(* IEC 61131-3 sources: plc-st-coding-agent/progress/evidence/f14_v14_remaining_20261113/jobs/codex_minimax-m27 (part 2) *)

(* ---- public-hard-01.raw_candidate_02.st ---- *)
FUNCTION_BLOCK MaterialProportioning
VAR_INPUT
    estop           : BOOL;          // Emergency stop signal (FALSE = stopped)
    opeMode         : BOOL;          // Operation mode (FALSE = manual, TRUE = automatic)
    valveAStart     : BOOL;          // Valve A start button
    valveBStart     : BOOL;          // Valve B start button
    valveCStart     : BOOL;          // Valve C start button
    valveDStart     : BOOL;          // Valve D start button
    mixMotorStart   : BOOL;          // Mixing motor start button
    autoStart       : BOOL;          // Automatic start button
    processMode     : BOOL;          // Process mode (FALSE = simple, TRUE = with C)
    levelSensor     : INT;           // Liquid level sensor (cm)
    mixMotorComplete: BOOL;          // Mixing complete signal
END_VAR
VAR_OUTPUT
    valveARun       : BOOL;          // Valve A run command
    valveBRun       : BOOL;          // Valve B run command
    valveCRun       : BOOL;          // Valve C run command
    valveDRun       : BOOL;          // Valve D run command
    mixMotorRun     : BOOL;          // Mixing motor run command
END_VAR
VAR
    // Rising edge detection for manual toggle buttons
    tmp_autoStart        : R_TRIG;
    tmp_valveAStart      : R_TRIG;
    tmp_valveBStart      : R_TRIG;
    tmp_valveCStart      : R_TRIG;
    tmp_valveDStart      : R_TRIG;
    tmp_mixMotorStart    : R_TRIG;

    // Automatic mode state machine
    tmp_autoState   : INT;           // 0=idle, 1=fillA, 2=fillB, 3=fillC, 4=mix, 5=drain, 6=done

    // Manual mode toggle states
    tmp_manualValveA    : BOOL;
    tmp_manualValveB    : BOOL;
    tmp_manualValveC    : BOOL;
    tmp_manualValveD    : BOOL;
    tmp_manualMixMotor  : BOOL;

    // Process complete flag for automatic mode
    tmp_autoComplete    : BOOL;
END_VAR

(* ENGINEERING_CONTRACT
================================================================================
Output          | Activation                  | Retention      | Reset
----------------|------------------------------|----------------|-------------------------
valveARun       | Manual: rising valveAStart   | Hold toggle    | estop, opeMode, auto step
                | Auto: state=1, level<50      |                |
PUB001, PUB002, PUB003, PUB004, PUB005, PUB006, PUB007, PUB008
----------------|------------------------------|----------------|-------------------------
valveBRun       | Auto: state=2, level<80      | Hold until 80cm| estop, opeMode, auto step
                |                              |                |
PUB003, PUB004, PUB006, PUB007, PUB008
----------------|------------------------------|----------------|-------------------------
valveCRun       | Auto: state=3, level<100     | Hold until 100cm| estop, opeMode, auto step
                | (processMode=true only)      |                |
PUB003, PUB004, PUB006, PUB007, PUB008
----------------|------------------------------|----------------|-------------------------
valveDRun       | Auto: mixMotorComplete       | Hold until reset| estop, opeMode, autoStart
                |                              |                |
PUB007, PUB008, PUB011, PUB012, PUB013, PUB014, PUB015
----------------|------------------------------|----------------|-------------------------
mixMotorRun     | Auto: state=4                | Hold until complete| estop, opeMode, autoStart
                | Manual: rising mixMotorStart |                |
PUB007, PUB008, PUB011, PUB012, PUB013, PUB014, PUB015
================================================================================
Priority: estop > manual/automatic mode switch > same-scan state updates
Boundary: levelSensor thresholds at 50cm, 80cm, 100cm (>= comparisons)
================================================================================
*)

(* CONTRACT_RULES [] *)

// Detect rising edges for toggle buttons
tmp_autoStart(CLK := autoStart);
tmp_valveAStart(CLK := valveAStart);
tmp_valveBStart(CLK := valveBStart);
tmp_valveCStart(CLK := valveCStart);
tmp_valveDStart(CLK := valveDStart);
tmp_mixMotorStart(CLK := mixMotorStart);

// Emergency stop: all equipment OFF immediately
IF NOT estop THEN
    valveARun := FALSE;
    valveBRun := FALSE;
    valveCRun := FALSE;
    valveDRun := FALSE;
    mixMotorRun := FALSE;
    tmp_autoState := 0;
    tmp_autoComplete := FALSE;
    tmp_manualValveA := FALSE;
    tmp_manualValveB := FALSE;
    tmp_manualValveC := FALSE;
    tmp_manualValveD := FALSE;
    tmp_manualMixMotor := FALSE;
    RETURN;
END_IF;

// Mode selection
IF opeMode THEN
    // AUTOMATIC MODE
    // Rising edge of autoStart initiates process
    IF tmp_autoStart.Q AND tmp_autoState = 0 THEN
        tmp_autoState := 1;
        tmp_autoComplete := FALSE;
    END_IF;

    // State machine execution
    CASE tmp_autoState OF
        0:  // Idle - all off
            valveARun := FALSE;
            valveBRun := FALSE;
            valveCRun := FALSE;
            valveDRun := FALSE;
            mixMotorRun := FALSE;

        1:  // Fill with valve A until level >= 50cm
            valveARun := TRUE;
            valveBRun := FALSE;
            valveCRun := FALSE;
            valveDRun := FALSE;
            mixMotorRun := FALSE;
            IF levelSensor >= 50 THEN
                valveARun := FALSE;
                tmp_autoState := 2;
            END_IF;

        2:  // Fill with valve B until level >= 80cm
            valveARun := FALSE;
            valveBRun := TRUE;
            valveCRun := FALSE;
            valveDRun := FALSE;
            mixMotorRun := FALSE;
            IF levelSensor >= 80 THEN
                valveBRun := FALSE;
                // Check processMode to determine next state
                IF processMode THEN
                    tmp_autoState := 3;  // Go to valve C
                ELSE
                    tmp_autoState := 4;  // Go directly to mixing
                END_IF;
            END_IF;

        3:  // Fill with valve C (processMode=true) until level >= 100cm
            valveARun := FALSE;
            valveBRun := FALSE;
            valveCRun := TRUE;
            valveDRun := FALSE;
            mixMotorRun := FALSE;
            IF levelSensor >= 100 THEN
                valveCRun := FALSE;
                tmp_autoState := 4;
            END_IF;

        4:  // Mixing until mixMotorComplete signal
            valveARun := FALSE;
            valveBRun := FALSE;
            valveCRun := FALSE;
            valveDRun := FALSE;
            mixMotorRun := TRUE;
            IF mixMotorComplete THEN
                mixMotorRun := FALSE;
                tmp_autoState := 5;
            END_IF;

        5:  // Open valve D to drain
            valveARun := FALSE;
            valveBRun := FALSE;
            valveCRun := FALSE;
            valveDRun := TRUE;
            mixMotorRun := FALSE;
            tmp_autoComplete := TRUE;
            tmp_autoState := 6;

        6:  // Process complete - valve D remains open until reset
            valveARun := FALSE;
            valveBRun := FALSE;
            valveCRun := FALSE;
            valveDRun := TRUE;
            mixMotorRun := FALSE;
            // Wait for autoStart to reset
            IF tmp_autoStart.Q THEN
                tmp_autoState := 0;
                tmp_autoComplete := FALSE;
            END_IF;
    END_CASE;

ELSE
    // MANUAL MODE
    // Reset automatic state when switching to manual
    tmp_autoState := 0;
    tmp_autoComplete := FALSE;

    // Toggle valve A
    IF tmp_valveAStart.Q THEN
        tmp_manualValveA := NOT tmp_manualValveA;
    END_IF;

    // Toggle valve B
    IF tmp_valveBStart.Q THEN
        tmp_manualValveB := NOT tmp_manualValveB;
    END_IF;

    // Toggle valve C
    IF tmp_valveCStart.Q THEN
        tmp_manualValveC := NOT tmp_manualValveC;
    END_IF;

    // Toggle valve D
    IF tmp_valveDStart.Q THEN
        tmp_manualValveD := NOT tmp_manualValveD;
    END_IF;

    // Toggle mixing motor
    IF tmp_mixMotorStart.Q THEN
        tmp_manualMixMotor := NOT tmp_manualMixMotor;
    END_IF;

    // Assign manual toggle states to outputs
    valveARun := tmp_manualValveA;
    valveBRun := tmp_manualValveB;
    valveCRun := tmp_manualValveC;
    valveDRun := tmp_manualValveD;
    mixMotorRun := tmp_manualMixMotor;
END_IF;

END_FUNCTION_BLOCK

(* ---- public-hard-02.candidate_01.st ---- *)
(* ENGINEERING_CONTRACT *)
(*
1. State Machine: IDLE | MOVING | PROCESSING | DONE
   - IDLE: Wait for sensor1 + station1Start to begin sequence
   - MOVING: Conveyor active, track position until sensor confirms arrival
   - PROCESSING: At processing station (2-4), wait for completion signal
   - DONE: At station 5, reset to IDLE next scan

2. Output Behavior:
   - conveyorLeft: Activated when targetStation < currentPosition (left movement)
   - conveyorRight: Activated when targetStation > currentPosition (right movement)
   - Both outputs OFF in IDLE, PROCESSING, and DONE states
   - Mutually exclusive per physical-direction rule (PUB001)

3. Retention:
   - currentPosition: Retains value between scans (product location)
   - sequenceIndex: Retains value between scans; resets to 1 on IDLE entry
   - Outputs: Default to FALSE on first scan

4. First Scan:
   - currentPosition := 1, sequenceIndex := 1
   - No conveyor movement until start conditions met

5. Explicit Reset:
   - DONE state: sequenceIndex := processLength + 1
   - Returns to IDLE next scan; sequenceIndex reset to 1 on new start

6. Same-Scan Priority:
   - Position update and conveyor enable use same-scan sensor values
   - Target station check confirms via sensor before stopping conveyor
   - No additional scan delay introduced

7. Units/Boundaries:
   - processLength: 1..8
   - currentPosition: 1..5 (station numbers)
   - sequenceIndex: 1..processLength+1
   - Stations: 1=loading, 2-4=processing, 5=output/storage
   - Station 5 has no completion signal (PUB003)
*)

(* CONTRACT_RULES [] *)

FUNCTION_BLOCK FlexibleProcessingControl
VAR_INPUT
    processLength : USINT := 8;
    sensor1 : BOOL;
    sensor2 : BOOL;
    sensor3 : BOOL;
    sensor4 : BOOL;
    sensor5 : BOOL;
    station1Start : BOOL;
    station2Complete : BOOL;
    station3Complete : BOOL;
    station4Complete : BOOL;
    processSequence : ARRAY[1..8] OF USINT;
END_VAR
VAR_OUTPUT
    conveyorLeft : BOOL;
    conveyorRight : BOOL;
END_VAR
VAR
    state : (IDLE, MOVING, PROCESSING, DONE) := IDLE;
    currentPosition : USINT := 1;
    sequenceIndex : USINT := 1;
    targetStation : USINT;
END_VAR

// Reset outputs by default
conveyorLeft := FALSE;
conveyorRight := FALSE;

// State machine implementation
CASE state OF
    IDLE:
        // Wait for material at station 1 and start button
        IF sensor1 AND station1Start THEN
            sequenceIndex := 1;
            targetStation := processSequence[sequenceIndex];
            sequenceIndex := sequenceIndex + 1;
            state := MOVING;
        END_IF;

    MOVING:
        // Determine conveyor direction and move toward target
        IF targetStation > currentPosition THEN
            currentPosition := currentPosition + 1;
            conveyorRight := TRUE;
            conveyorLeft := FALSE;
        ELSIF targetStation < currentPosition THEN
            currentPosition := currentPosition - 1;
            conveyorLeft := TRUE;
            conveyorRight := FALSE;
        END_IF;

        // Check if product reached target station via sensor confirmation
        IF currentPosition = targetStation THEN
            // Verify arrival with appropriate sensor
            IF (currentPosition = 1 AND sensor1) OR
               (currentPosition = 2 AND sensor2) OR
               (currentPosition = 3 AND sensor3) OR
               (currentPosition = 4 AND sensor4) OR
               (currentPosition = 5 AND sensor5) THEN
                conveyorLeft := FALSE;
                conveyorRight := FALSE;

                // Station 5 is output/storage - no completion signal
                IF currentPosition = 5 THEN
                    state := DONE;
                ELSE
                    state := PROCESSING;
                END_IF;
            END_IF;
        END_IF;

    PROCESSING:
        // Wait for processing completion at stations 2-4
        IF (currentPosition = 2 AND station2Complete) OR
           (currentPosition = 3 AND station3Complete) OR
           (currentPosition = 4 AND station4Complete) THEN
            // Check if next target is station 5 (final output)
            IF targetStation = 5 THEN
                state := DONE;
            ELSIF sequenceIndex <= processLength THEN
                targetStation := processSequence[sequenceIndex];
                sequenceIndex := sequenceIndex + 1;
                state := MOVING;
            ELSE
                // Sequence complete, product should be at station 5
                state := DONE;
            END_IF;
        END_IF;

    DONE:
        // Product reached station 5, prepare for next cycle
        sequenceIndex := processLength + 1;
        state := IDLE;
END_CASE;
END_FUNCTION_BLOCK

(* ---- public-hard-02.raw_candidate_01.st ---- *)
(* ENGINEERING_CONTRACT *)
(*
1. State Machine: IDLE | MOVING | PROCESSING | DONE
   - IDLE: Wait for sensor1 + station1Start to begin sequence
   - MOVING: Conveyor active, track position until sensor confirms arrival
   - PROCESSING: At processing station (2-4), wait for completion signal
   - DONE: At station 5, reset to IDLE next scan

2. Output Behavior:
   - conveyorLeft: Activated when targetStation < currentPosition (left movement)
   - conveyorRight: Activated when targetStation > currentPosition (right movement)
   - Both outputs OFF in IDLE, PROCESSING, and DONE states
   - Mutually exclusive per physical-direction rule (PUB001)

3. Retention:
   - currentPosition: Retains value between scans (product location)
   - sequenceIndex: Retains value between scans; resets to 1 on IDLE entry
   - Outputs: Default to FALSE on first scan

4. First Scan:
   - currentPosition := 1, sequenceIndex := 1
   - No conveyor movement until start conditions met

5. Explicit Reset:
   - DONE state: sequenceIndex := processLength + 1
   - Returns to IDLE next scan; sequenceIndex reset to 1 on new start

6. Same-Scan Priority:
   - Position update and conveyor enable use same-scan sensor values
   - Target station check confirms via sensor before stopping conveyor
   - No additional scan delay introduced

7. Units/Boundaries:
   - processLength: 1..8
   - currentPosition: 1..5 (station numbers)
   - sequenceIndex: 1..processLength+1
   - Stations: 1=loading, 2-4=processing, 5=output/storage
   - Station 5 has no completion signal (PUB003)
*)

(* CONTRACT_RULES [] *)

FUNCTION_BLOCK FlexibleProcessingControl
VAR_INPUT
    processLength : USINT := 8;
    sensor1 : BOOL;
    sensor2 : BOOL;
    sensor3 : BOOL;
    sensor4 : BOOL;
    sensor5 : BOOL;
    station1Start : BOOL;
    station2Complete : BOOL;
    station3Complete : BOOL;
    station4Complete : BOOL;
    processSequence : ARRAY[1..8] OF USINT;
END_VAR
VAR_OUTPUT
    conveyorLeft : BOOL;
    conveyorRight : BOOL;
END_VAR
VAR
    state : (IDLE, MOVING, PROCESSING, DONE) := IDLE;
    currentPosition : USINT := 1;
    sequenceIndex : USINT := 1;
    targetStation : USINT;
END_VAR

// Reset outputs by default
conveyorLeft := FALSE;
conveyorRight := FALSE;

// State machine implementation
CASE state OF
    IDLE:
        // Wait for material at station 1 and start button
        IF sensor1 AND station1Start THEN
            sequenceIndex := 1;
            targetStation := processSequence[sequenceIndex];
            sequenceIndex := sequenceIndex + 1;
            state := MOVING;
        END_IF;

    MOVING:
        // Determine conveyor direction and move toward target
        IF targetStation > currentPosition THEN
            currentPosition := currentPosition + 1;
            conveyorRight := TRUE;
            conveyorLeft := FALSE;
        ELSIF targetStation < currentPosition THEN
            currentPosition := currentPosition - 1;
            conveyorLeft := TRUE;
            conveyorRight := FALSE;
        END_IF;

        // Check if product reached target station via sensor confirmation
        IF currentPosition = targetStation THEN
            // Verify arrival with appropriate sensor
            IF (currentPosition = 1 AND sensor1) OR
               (currentPosition = 2 AND sensor2) OR
               (currentPosition = 3 AND sensor3) OR
               (currentPosition = 4 AND sensor4) OR
               (currentPosition = 5 AND sensor5) THEN
                conveyorLeft := FALSE;
                conveyorRight := FALSE;

                // Station 5 is output/storage - no completion signal
                IF currentPosition = 5 THEN
                    state := DONE;
                ELSE
                    state := PROCESSING;
                END_IF;
            END_IF;
        END_IF;

    PROCESSING:
        // Wait for processing completion at stations 2-4
        IF (currentPosition = 2 AND station2Complete) OR
           (currentPosition = 3 AND station3Complete) OR
           (currentPosition = 4 AND station4Complete) THEN
            // Check if next target is station 5 (final output)
            IF targetStation = 5 THEN
                state := DONE;
            ELSIF sequenceIndex <= processLength THEN
                targetStation := processSequence[sequenceIndex];
                sequenceIndex := sequenceIndex + 1;
                state := MOVING;
            ELSE
                // Sequence complete, product should be at station 5
                state := DONE;
            END_IF;
        END_IF;

    DONE:
        // Product reached station 5, prepare for next cycle
        sequenceIndex := processLength + 1;
        state := IDLE;
END_CASE;
END_FUNCTION_BLOCK

(* ---- public-hard-03.candidate_01.st ---- *)
(* ENGINEERING_CONTRACT *)
(*
  Operation Priority (PUB001): Sequential evaluation order
    1. QUERY   - Read-only, sets recipeQueryResult
    2. ADD     - Write to empty slot, sets recipeAdded
    3. DELETE  - Write-clear slot, sets recipeDeleted
    4. MODIFY  - Write-replace slot, sets recipeModified

  Activation  : Edge-triggered via R_TRIG on command inputs
  Retention   : All outputs (except recipeQueryResult) are single-scan pulses
  Reset       : Outputs clear on subsequent scans when command deasserted
  Same-scan   : Final command state determines which R_TRIG fires
  Error       : error=TRUE with status code, no data written
  Success     : Specific success flag TRUE, error=FALSE, status=0
*)

(* CONTRACT_RULES [] *)

FUNCTION_BLOCK RecipeManagement
VAR_INPUT
    addRecipe    : BOOL;
    deleteRecipe : BOOL;
    modifyRecipe : BOOL;
    queryRecipe  : BOOL;
    recipeIn     : ST_Recipe;
END_VAR

VAR_OUTPUT
    recipeAdded       : BOOL := FALSE;
    recipeDeleted     : BOOL := FALSE;
    recipeModified    : BOOL := FALSE;
    recipeQueryResult : ST_Recipe;
    error             : BOOL := FALSE;
    status            : WORD := 0;
END_VAR

VAR_IN_OUT
    recipe : ARRAY[1..10] OF ST_Recipe;
END_VAR

VAR
    trigAdd    : R_TRIG;
    trigDelete : R_TRIG;
    trigModify : R_TRIG;
    trigQuery  : R_TRIG;
    tmp_i      : INT;
    tmp_slot   : INT;
    tmp_found  : BOOL;
    tmp_empty  : BOOL;
END_VAR

// Clear output flags at start of each scan
recipeAdded    := FALSE;
recipeDeleted  := FALSE;
recipeModified := FALSE;
error          := FALSE;
status         := 0;

// Detect rising edges on command inputs
trigQuery(IN:=queryRecipe);
trigAdd(IN:=addRecipe);
trigDelete(IN:=deleteRecipe);
trigModify(IN:=modifyRecipe);

// Operation 1: Query Recipe (PUB002, PUB008)
IF trigQuery.Q THEN
    tmp_found := FALSE;
    tmp_i := 1;
    WHILE tmp_i <= 10 AND NOT tmp_found DO
        IF recipe[tmp_i].recipeID = recipeIn.recipeID THEN
            tmp_found := TRUE;
        ELSE
            tmp_i := tmp_i + 1;
        END_IF;
    END_WHILE;

    IF tmp_found THEN
        recipeQueryResult := recipe[tmp_i];
        error   := FALSE;
        status  := 0;
    ELSE
        error   := TRUE;
        status  := 16#8001;  // Recipe not found
    END_IF;
END_IF;

// Operation 2: Add Recipe (PUB003, PUB009)
IF trigAdd.Q THEN
    // Check for duplicate recipeID
    tmp_found := FALSE;
    tmp_i := 1;
    WHILE tmp_i <= 10 AND NOT tmp_found DO
        IF recipe[tmp_i].recipeID = recipeIn.recipeID THEN
            tmp_found := TRUE;
        ELSE
            tmp_i := tmp_i + 1;
        END_IF;
    END_WHILE;

    IF tmp_found THEN
        error   := TRUE;
        status  := 16#8002;  // Duplicate recipeID
    ELSE
        // Find first empty slot (smallest index)
        tmp_empty := FALSE;
        tmp_slot  := 1;
        WHILE tmp_slot <= 10 AND NOT tmp_empty DO
            IF recipe[tmp_slot].recipeID = 0 THEN
                tmp_empty := TRUE;
            ELSE
                tmp_slot := tmp_slot + 1;
            END_IF;
        END_WHILE;

        IF tmp_empty THEN
            recipe[tmp_slot] := recipeIn;
            recipeAdded := TRUE;
            error       := FALSE;
            status      := 0;
        ELSE
            error   := TRUE;
            status  := 16#8003;  // No empty slot
        END_IF;
    END_IF;
END_IF;

// Operation 3: Delete Recipe (PUB004, PUB010)
IF trigDelete.Q THEN
    tmp_found := FALSE;
    tmp_i := 1;
    WHILE tmp_i <= 10 AND NOT tmp_found DO
        IF recipe[tmp_i].recipeID = recipeIn.recipeID THEN
            tmp_found := TRUE;
        ELSE
            tmp_i := tmp_i + 1;
        END_IF;
    END_WHILE;

    IF tmp_found THEN
        recipe[tmp_i].recipeID         := 0;
        recipe[tmp_i].ingredientType   := 0;
        recipe[tmp_i].ingredientRatio  := 0.0;
        recipe[tmp_i].productionTemperature := 0.0;
        recipeDeleted := TRUE;
        error         := FALSE;
        status        := 0;
    ELSE
        error   := TRUE;
        status  := 16#8004;  // Recipe not found for deletion
    END_IF;
END_IF;

// Operation 4: Modify Recipe (PUB005, PUB011)
IF trigModify.Q THEN
    tmp_found := FALSE;
    tmp_i := 1;
    WHILE tmp_i <= 10 AND NOT tmp_found DO
        IF recipe[tmp_i].recipeID = recipeIn.recipeID THEN
            tmp_found := TRUE;
        ELSE
            tmp_i := tmp_i + 1;
        END_IF;
    END_WHILE;

    IF tmp_found THEN
        recipe[tmp_i] := recipeIn;
        recipeModified := TRUE;
        error          := FALSE;
        status         := 0;
    ELSE
        error   := TRUE;
        status  := 16#8005;  // Recipe not found for modification
    END_IF;
END_IF;

END_FUNCTION_BLOCK

(* ---- public-hard-03.candidate_02.st ---- *)
(* ENGINEERING_CONTRACT *)
(*
  Operation Priority (PUB001): Sequential evaluation order
    1. QUERY   - Read-only, sets recipeQueryResult
    2. ADD     - Write to empty slot, sets recipeAdded
    3. DELETE  - Write-clear slot, sets recipeDeleted
    4. MODIFY  - Write-replace slot, sets recipeModified

  Activation  : Edge-triggered via R_TRIG on command inputs
  Retention   : All outputs (except recipeQueryResult) are single-scan pulses
  Reset       : Outputs clear on subsequent scans when command deasserted
  Same-scan   : Final command state determines which R_TRIG fires
  Error       : error=TRUE with status code, no data written
  Success     : Specific success flag TRUE, error=FALSE, status=0
*)

TYPE ST_Recipe : STRUCT
    recipeID              : INT;
    ingredientType        : INT;
    ingredientRatio       : REAL;
    productionTemperature : REAL;
END_STRUCT END_TYPE;

(* CONTRACT_RULES [] *)

FUNCTION_BLOCK RecipeManagement
VAR_INPUT
    addRecipe    : BOOL;
    deleteRecipe : BOOL;
    modifyRecipe : BOOL;
    queryRecipe  : BOOL;
    recipeIn     : ST_Recipe;
END_VAR

VAR_OUTPUT
    recipeAdded       : BOOL := FALSE;
    recipeDeleted     : BOOL := FALSE;
    recipeModified    : BOOL := FALSE;
    recipeQueryResult : ST_Recipe;
    error             : BOOL := FALSE;
    status            : WORD := 0;
END_VAR

VAR_IN_OUT
    recipe : ARRAY[1..10] OF ST_Recipe;
END_VAR

VAR
    trigAdd    : R_TRIG;
    trigDelete : R_TRIG;
    trigModify : R_TRIG;
    trigQuery  : R_TRIG;
    tmp_i      : INT;
    tmp_slot   : INT;
    tmp_found  : BOOL;
    tmp_empty  : BOOL;
END_VAR

// Clear output flags at start of each scan
recipeAdded    := FALSE;
recipeDeleted  := FALSE;
recipeModified := FALSE;
error          := FALSE;
status         := 0;

// Detect rising edges on command inputs
trigQuery(CLK:=queryRecipe);
trigAdd(CLK:=addRecipe);
trigDelete(CLK:=deleteRecipe);
trigModify(CLK:=modifyRecipe);

// Operation 1: Query Recipe (PUB002, PUB008)
IF trigQuery.Q THEN
    tmp_found := FALSE;
    tmp_i := 1;
    WHILE tmp_i <= 10 AND NOT tmp_found DO
        IF recipe[tmp_i].recipeID = recipeIn.recipeID THEN
            tmp_found := TRUE;
        ELSE
            tmp_i := tmp_i + 1;
        END_IF;
    END_WHILE;

    IF tmp_found THEN
        recipeQueryResult := recipe[tmp_i];
        error   := FALSE;
        status  := 0;
    ELSE
        error   := TRUE;
        status  := 16#8001;  // Recipe not found
    END_IF;
END_IF;

// Operation 2: Add Recipe (PUB003, PUB009)
IF trigAdd.Q THEN
    // Check for duplicate recipeID
    tmp_found := FALSE;
    tmp_i := 1;
    WHILE tmp_i <= 10 AND NOT tmp_found DO
        IF recipe[tmp_i].recipeID = recipeIn.recipeID THEN
            tmp_found := TRUE;
        ELSE
            tmp_i := tmp_i + 1;
        END_IF;
    END_WHILE;

    IF tmp_found THEN
        error   := TRUE;
        status  := 16#8002;  // Duplicate recipeID
    ELSE
        // Find first empty slot (smallest index)
        tmp_empty := FALSE;
        tmp_slot  := 1;
        WHILE tmp_slot <= 10 AND NOT tmp_empty DO
            IF recipe[tmp_slot].recipeID = 0 THEN
                tmp_empty := TRUE;
            ELSE
                tmp_slot := tmp_slot + 1;
            END_IF;
        END_WHILE;

        IF tmp_empty THEN
            recipe[tmp_slot] := recipeIn;
            recipeAdded := TRUE;
            error       := FALSE;
            status      := 0;
        ELSE
            error   := TRUE;
            status  := 16#8003;  // No empty slot
        END_IF;
    END_IF;
END_IF;

// Operation 3: Delete Recipe (PUB004, PUB010)
IF trigDelete.Q THEN
    tmp_found := FALSE;
    tmp_i := 1;
    WHILE tmp_i <= 10 AND NOT tmp_found DO
        IF recipe[tmp_i].recipeID = recipeIn.recipeID THEN
            tmp_found := TRUE;
        ELSE
            tmp_i := tmp_i + 1;
        END_IF;
    END_WHILE;

    IF tmp_found THEN
        recipe[tmp_i].recipeID         := 0;
        recipe[tmp_i].ingredientType   := 0;
        recipe[tmp_i].ingredientRatio  := 0.0;
        recipe[tmp_i].productionTemperature := 0.0;
        recipeDeleted := TRUE;
        error         := FALSE;
        status        := 0;
    ELSE
        error   := TRUE;
        status  := 16#8004;  // Recipe not found for deletion
    END_IF;
END_IF;

// Operation 4: Modify Recipe (PUB005, PUB011)
IF trigModify.Q THEN
    tmp_found := FALSE;
    tmp_i := 1;
    WHILE tmp_i <= 10 AND NOT tmp_found DO
        IF recipe[tmp_i].recipeID = recipeIn.recipeID THEN
            tmp_found := TRUE;
        ELSE
            tmp_i := tmp_i + 1;
        END_IF;
    END_WHILE;

    IF tmp_found THEN
        recipe[tmp_i] := recipeIn;
        recipeModified := TRUE;
        error          := FALSE;
        status         := 0;
    ELSE
        error   := TRUE;
        status  := 16#8005;  // Recipe not found for modification
    END_IF;
END_IF;

END_FUNCTION_BLOCK

(* ---- public-hard-03.candidate_04.st ---- *)
(* ENGINEERING_CONTRACT *)
(*
  Operation Priority (PUB001): Sequential evaluation order
    1. QUERY   - Read-only, sets recipeQueryResult
    2. ADD     - Write to empty slot, sets recipeAdded
    3. DELETE  - Write-clear slot, sets recipeDeleted
    4. MODIFY  - Write-replace slot, sets recipeModified

  Activation  : Edge-triggered via R_TRIG on command inputs
  Retention   : All outputs (except recipeQueryResult) are single-scan pulses
  Reset       : Outputs clear on subsequent scans when command deasserted
  Same-scan   : Final command state determines which R_TRIG fires
  Error       : error=TRUE with status code, no data written
  Success     : Specific success flag TRUE, error=FALSE, status=0
*)

TYPE ST_Recipe : STRUCT
    recipeID              : INT;
    ingredientType        : INT;
    ingredientRatio       : REAL;
    productionTemperature : REAL;
END_STRUCT END_TYPE;

(* CONTRACT_RULES [] *)

FUNCTION_BLOCK RecipeManagement
VAR_INPUT
    addRecipe    : BOOL;
    deleteRecipe : BOOL;
    modifyRecipe : BOOL;
    queryRecipe  : BOOL;
    recipeIn     : ST_Recipe;
END_VAR

VAR_OUTPUT
    recipeAdded       : BOOL := FALSE;
    recipeDeleted     : BOOL := FALSE;
    recipeModified    : BOOL := FALSE;
    recipeQueryResult : ST_Recipe;
    error             : BOOL := FALSE;
    status            : WORD := 0;
END_VAR

VAR_IN_OUT
    recipe : ARRAY[1..10] OF ST_Recipe;
END_VAR

VAR
    trigAdd    : R_TRIG;
    trigDelete : R_TRIG;
    trigModify : R_TRIG;
    trigQuery  : R_TRIG;
    tmp_i      : INT;
    tmp_slot   : INT;
    tmp_found  : BOOL;
    tmp_empty  : BOOL;
END_VAR

// Clear output flags at start of each scan
recipeAdded    := FALSE;
recipeDeleted  := FALSE;
recipeModified := FALSE;
IF trigQuery.Q OR trigAdd.Q OR trigDelete.Q OR trigModify.Q THEN
    error   := FALSE;
    status  := 0;
END_IF;

// Detect rising edges on command inputs
trigQuery(CLK:=queryRecipe);
trigAdd(CLK:=addRecipe);
trigDelete(CLK:=deleteRecipe);
trigModify(CLK:=modifyRecipe);

// Operation 1: Query Recipe (PUB002, PUB008)
IF trigQuery.Q THEN
    tmp_found := FALSE;
    tmp_i := 1;
    WHILE tmp_i <= 10 AND NOT tmp_found DO
        IF recipe[tmp_i].recipeID = recipeIn.recipeID THEN
            tmp_found := TRUE;
        ELSE
            tmp_i := tmp_i + 1;
        END_IF;
    END_WHILE;

    IF tmp_found THEN
        recipeQueryResult := recipe[tmp_i];
        error   := FALSE;
        status  := 0;
    ELSE
        error   := TRUE;
        status  := 16#8001;  // Recipe not found
    END_IF;
END_IF;

// Operation 2: Add Recipe (PUB003, PUB009)
IF trigAdd.Q THEN
    // Check for duplicate recipeID
    tmp_found := FALSE;
    tmp_i := 1;
    WHILE tmp_i <= 10 AND NOT tmp_found DO
        IF recipe[tmp_i].recipeID = recipeIn.recipeID THEN
            tmp_found := TRUE;
        ELSE
            tmp_i := tmp_i + 1;
        END_IF;
    END_WHILE;

    IF tmp_found THEN
        error   := TRUE;
        status  := 16#8002;  // Duplicate recipeID
    ELSE
        // Find first empty slot (smallest index)
        tmp_empty := FALSE;
        tmp_slot  := 1;
        WHILE tmp_slot <= 10 AND NOT tmp_empty DO
            IF recipe[tmp_slot].recipeID = 0 THEN
                tmp_empty := TRUE;
            ELSE
                tmp_slot := tmp_slot + 1;
            END_IF;
        END_WHILE;

        IF tmp_empty THEN
            recipe[tmp_slot] := recipeIn;
            recipeAdded := TRUE;
            error       := FALSE;
            status      := 0;
        ELSE
            error   := TRUE;
            status  := 16#8003;  // No empty slot
        END_IF;
    END_IF;
END_IF;

// Operation 3: Delete Recipe (PUB004, PUB010)
IF trigDelete.Q THEN
    tmp_found := FALSE;
    tmp_i := 1;
    WHILE tmp_i <= 10 AND NOT tmp_found DO
        IF recipe[tmp_i].recipeID = recipeIn.recipeID THEN
            tmp_found := TRUE;
        ELSE
            tmp_i := tmp_i + 1;
        END_IF;
    END_WHILE;

    IF tmp_found THEN
        recipe[tmp_i].recipeID         := 0;
        recipe[tmp_i].ingredientType   := 0;
        recipe[tmp_i].ingredientRatio  := 0.0;
        recipe[tmp_i].productionTemperature := 0.0;
        recipeDeleted := TRUE;
        error         := FALSE;
        status        := 0;
    ELSE
        error   := TRUE;
        status  := 16#8004;  // Recipe not found for deletion
    END_IF;
END_IF;

// Operation 4: Modify Recipe (PUB005, PUB011)
IF trigModify.Q THEN
    tmp_found := FALSE;
    tmp_i := 1;
    WHILE tmp_i <= 10 AND NOT tmp_found DO
        IF recipe[tmp_i].recipeID = recipeIn.recipeID THEN
            tmp_found := TRUE;
        ELSE
            tmp_i := tmp_i + 1;
        END_IF;
    END_WHILE;

    IF tmp_found THEN
        recipe[tmp_i] := recipeIn;
        recipeModified := TRUE;
        error          := FALSE;
        status         := 0;
    ELSE
        error   := TRUE;
        status  := 16#8005;  // Recipe not found for modification
    END_IF;
END_IF;

END_FUNCTION_BLOCK

(* ---- public-hard-03.patch_base_02.st ---- *)
(* ENGINEERING_CONTRACT *)
(*
  Operation Priority (PUB001): Sequential evaluation order
    1. QUERY   - Read-only, sets recipeQueryResult
    2. ADD     - Write to empty slot, sets recipeAdded
    3. DELETE  - Write-clear slot, sets recipeDeleted
    4. MODIFY  - Write-replace slot, sets recipeModified

  Activation  : Edge-triggered via R_TRIG on command inputs
  Retention   : All outputs (except recipeQueryResult) are single-scan pulses
  Reset       : Outputs clear on subsequent scans when command deasserted
  Same-scan   : Final command state determines which R_TRIG fires
  Error       : error=TRUE with status code, no data written
  Success     : Specific success flag TRUE, error=FALSE, status=0
*)

(* CONTRACT_RULES [] *)

FUNCTION_BLOCK RecipeManagement
VAR_INPUT
    addRecipe    : BOOL;
    deleteRecipe : BOOL;
    modifyRecipe : BOOL;
    queryRecipe  : BOOL;
    recipeIn     : ST_Recipe;
END_VAR

VAR_OUTPUT
    recipeAdded       : BOOL := FALSE;
    recipeDeleted     : BOOL := FALSE;
    recipeModified    : BOOL := FALSE;
    recipeQueryResult : ST_Recipe;
    error             : BOOL := FALSE;
    status            : WORD := 0;
END_VAR

VAR_IN_OUT
    recipe : ARRAY[1..10] OF ST_Recipe;
END_VAR

VAR
    trigAdd    : R_TRIG;
    trigDelete : R_TRIG;
    trigModify : R_TRIG;
    trigQuery  : R_TRIG;
    tmp_i      : INT;
    tmp_slot   : INT;
    tmp_found  : BOOL;
    tmp_empty  : BOOL;
END_VAR

// Clear output flags at start of each scan
recipeAdded    := FALSE;
recipeDeleted  := FALSE;
recipeModified := FALSE;
error          := FALSE;
status         := 0;

// Detect rising edges on command inputs
trigQuery(IN:=queryRecipe);
trigAdd(IN:=addRecipe);
trigDelete(IN:=deleteRecipe);
trigModify(IN:=modifyRecipe);

// Operation 1: Query Recipe (PUB002, PUB008)
IF trigQuery.Q THEN
    tmp_found := FALSE;
    tmp_i := 1;
    WHILE tmp_i <= 10 AND NOT tmp_found DO
        IF recipe[tmp_i].recipeID = recipeIn.recipeID THEN
            tmp_found := TRUE;
        ELSE
            tmp_i := tmp_i + 1;
        END_IF;
    END_WHILE;

    IF tmp_found THEN
        recipeQueryResult := recipe[tmp_i];
        error   := FALSE;
        status  := 0;
    ELSE
        error   := TRUE;
        status  := 16#8001;  // Recipe not found
    END_IF;
END_IF;

// Operation 2: Add Recipe (PUB003, PUB009)
IF trigAdd.Q THEN
    // Check for duplicate recipeID
    tmp_found := FALSE;
    tmp_i := 1;
    WHILE tmp_i <= 10 AND NOT tmp_found DO
        IF recipe[tmp_i].recipeID = recipeIn.recipeID THEN
            tmp_found := TRUE;
        ELSE
            tmp_i := tmp_i + 1;
        END_IF;
    END_WHILE;

    IF tmp_found THEN
        error   := TRUE;
        status  := 16#8002;  // Duplicate recipeID
    ELSE
        // Find first empty slot (smallest index)
        tmp_empty := FALSE;
        tmp_slot  := 1;
        WHILE tmp_slot <= 10 AND NOT tmp_empty DO
            IF recipe[tmp_slot].recipeID = 0 THEN
                tmp_empty := TRUE;
            ELSE
                tmp_slot := tmp_slot + 1;
            END_IF;
        END_WHILE;

        IF tmp_empty THEN
            recipe[tmp_slot] := recipeIn;
            recipeAdded := TRUE;
            error       := FALSE;
            status      := 0;
        ELSE
            error   := TRUE;
            status  := 16#8003;  // No empty slot
        END_IF;
    END_IF;
END_IF;

// Operation 3: Delete Recipe (PUB004, PUB010)
IF trigDelete.Q THEN
    tmp_found := FALSE;
    tmp_i := 1;
    WHILE tmp_i <= 10 AND NOT tmp_found DO
        IF recipe[tmp_i].recipeID = recipeIn.recipeID THEN
            tmp_found := TRUE;
        ELSE
            tmp_i := tmp_i + 1;
        END_IF;
    END_WHILE;

    IF tmp_found THEN
        recipe[tmp_i].recipeID         := 0;
        recipe[tmp_i].ingredientType   := 0;
        recipe[tmp_i].ingredientRatio  := 0.0;
        recipe[tmp_i].productionTemperature := 0.0;
        recipeDeleted := TRUE;
        error         := FALSE;
        status        := 0;
    ELSE
        error   := TRUE;
        status  := 16#8004;  // Recipe not found for deletion
    END_IF;
END_IF;

// Operation 4: Modify Recipe (PUB005, PUB011)
IF trigModify.Q THEN
    tmp_found := FALSE;
    tmp_i := 1;
    WHILE tmp_i <= 10 AND NOT tmp_found DO
        IF recipe[tmp_i].recipeID = recipeIn.recipeID THEN
            tmp_found := TRUE;
        ELSE
            tmp_i := tmp_i + 1;
        END_IF;
    END_WHILE;

    IF tmp_found THEN
        recipe[tmp_i] := recipeIn;
        recipeModified := TRUE;
        error          := FALSE;
        status         := 0;
    ELSE
        error   := TRUE;
        status  := 16#8005;  // Recipe not found for modification
    END_IF;
END_IF;

END_FUNCTION_BLOCK

(* ---- public-hard-03.patch_base_03.st ---- *)
(* ENGINEERING_CONTRACT *)
(*
  Operation Priority (PUB001): Sequential evaluation order
    1. QUERY   - Read-only, sets recipeQueryResult
    2. ADD     - Write to empty slot, sets recipeAdded
    3. DELETE  - Write-clear slot, sets recipeDeleted
    4. MODIFY  - Write-replace slot, sets recipeModified

  Activation  : Edge-triggered via R_TRIG on command inputs
  Retention   : All outputs (except recipeQueryResult) are single-scan pulses
  Reset       : Outputs clear on subsequent scans when command deasserted
  Same-scan   : Final command state determines which R_TRIG fires
  Error       : error=TRUE with status code, no data written
  Success     : Specific success flag TRUE, error=FALSE, status=0
*)

TYPE ST_Recipe : STRUCT
    recipeID              : INT;
    ingredientType        : INT;
    ingredientRatio       : REAL;
    productionTemperature : REAL;
END_STRUCT END_TYPE;

(* CONTRACT_RULES [] *)

FUNCTION_BLOCK RecipeManagement
VAR_INPUT
    addRecipe    : BOOL;
    deleteRecipe : BOOL;
    modifyRecipe : BOOL;
    queryRecipe  : BOOL;
    recipeIn     : ST_Recipe;
END_VAR

VAR_OUTPUT
    recipeAdded       : BOOL := FALSE;
    recipeDeleted     : BOOL := FALSE;
    recipeModified    : BOOL := FALSE;
    recipeQueryResult : ST_Recipe;
    error             : BOOL := FALSE;
    status            : WORD := 0;
END_VAR

VAR_IN_OUT
    recipe : ARRAY[1..10] OF ST_Recipe;
END_VAR

VAR
    trigAdd    : R_TRIG;
    trigDelete : R_TRIG;
    trigModify : R_TRIG;
    trigQuery  : R_TRIG;
    tmp_i      : INT;
    tmp_slot   : INT;
    tmp_found  : BOOL;
    tmp_empty  : BOOL;
END_VAR

// Clear output flags at start of each scan
recipeAdded    := FALSE;
recipeDeleted  := FALSE;
recipeModified := FALSE;
error          := FALSE;
status         := 0;

// Detect rising edges on command inputs
trigQuery(CLK:=queryRecipe);
trigAdd(CLK:=addRecipe);
trigDelete(CLK:=deleteRecipe);
trigModify(CLK:=modifyRecipe);

// Operation 1: Query Recipe (PUB002, PUB008)
IF trigQuery.Q THEN
    tmp_found := FALSE;
    tmp_i := 1;
    WHILE tmp_i <= 10 AND NOT tmp_found DO
        IF recipe[tmp_i].recipeID = recipeIn.recipeID THEN
            tmp_found := TRUE;
        ELSE
            tmp_i := tmp_i + 1;
        END_IF;
    END_WHILE;

    IF tmp_found THEN
        recipeQueryResult := recipe[tmp_i];
        error   := FALSE;
        status  := 0;
    ELSE
        error   := TRUE;
        status  := 16#8001;  // Recipe not found
    END_IF;
END_IF;

// Operation 2: Add Recipe (PUB003, PUB009)
IF trigAdd.Q THEN
    // Check for duplicate recipeID
    tmp_found := FALSE;
    tmp_i := 1;
    WHILE tmp_i <= 10 AND NOT tmp_found DO
        IF recipe[tmp_i].recipeID = recipeIn.recipeID THEN
            tmp_found := TRUE;
        ELSE
            tmp_i := tmp_i + 1;
        END_IF;
    END_WHILE;

    IF tmp_found THEN
        error   := TRUE;
        status  := 16#8002;  // Duplicate recipeID
    ELSE
        // Find first empty slot (smallest index)
        tmp_empty := FALSE;
        tmp_slot  := 1;
        WHILE tmp_slot <= 10 AND NOT tmp_empty DO
            IF recipe[tmp_slot].recipeID = 0 THEN
                tmp_empty := TRUE;
            ELSE
                tmp_slot := tmp_slot + 1;
            END_IF;
        END_WHILE;

        IF tmp_empty THEN
            recipe[tmp_slot] := recipeIn;
            recipeAdded := TRUE;
            error       := FALSE;
            status      := 0;
        ELSE
            error   := TRUE;
            status  := 16#8003;  // No empty slot
        END_IF;
    END_IF;
END_IF;

// Operation 3: Delete Recipe (PUB004, PUB010)
IF trigDelete.Q THEN
    tmp_found := FALSE;
    tmp_i := 1;
    WHILE tmp_i <= 10 AND NOT tmp_found DO
        IF recipe[tmp_i].recipeID = recipeIn.recipeID THEN
            tmp_found := TRUE;
        ELSE
            tmp_i := tmp_i + 1;
        END_IF;
    END_WHILE;

    IF tmp_found THEN
        recipe[tmp_i].recipeID         := 0;
        recipe[tmp_i].ingredientType   := 0;
        recipe[tmp_i].ingredientRatio  := 0.0;
        recipe[tmp_i].productionTemperature := 0.0;
        recipeDeleted := TRUE;
        error         := FALSE;
        status        := 0;
    ELSE
        error   := TRUE;
        status  := 16#8004;  // Recipe not found for deletion
    END_IF;
END_IF;

// Operation 4: Modify Recipe (PUB005, PUB011)
IF trigModify.Q THEN
    tmp_found := FALSE;
    tmp_i := 1;
    WHILE tmp_i <= 10 AND NOT tmp_found DO
        IF recipe[tmp_i].recipeID = recipeIn.recipeID THEN
            tmp_found := TRUE;
        ELSE
            tmp_i := tmp_i + 1;
        END_IF;
    END_WHILE;

    IF tmp_found THEN
        recipe[tmp_i] := recipeIn;
        recipeModified := TRUE;
        error          := FALSE;
        status         := 0;
    ELSE
        error   := TRUE;
        status  := 16#8005;  // Recipe not found for modification
    END_IF;
END_IF;

END_FUNCTION_BLOCK

(* ---- public-hard-03.patch_base_04.st ---- *)
(* ENGINEERING_CONTRACT *)
(*
  Operation Priority (PUB001): Sequential evaluation order
    1. QUERY   - Read-only, sets recipeQueryResult
    2. ADD     - Write to empty slot, sets recipeAdded
    3. DELETE  - Write-clear slot, sets recipeDeleted
    4. MODIFY  - Write-replace slot, sets recipeModified

  Activation  : Edge-triggered via R_TRIG on command inputs
  Retention   : All outputs (except recipeQueryResult) are single-scan pulses
  Reset       : Outputs clear on subsequent scans when command deasserted
  Same-scan   : Final command state determines which R_TRIG fires
  Error       : error=TRUE with status code, no data written
  Success     : Specific success flag TRUE, error=FALSE, status=0
*)

TYPE ST_Recipe : STRUCT
    recipeID              : INT;
    ingredientType        : INT;
    ingredientRatio       : REAL;
    productionTemperature : REAL;
END_STRUCT END_TYPE;

(* CONTRACT_RULES [] *)

FUNCTION_BLOCK RecipeManagement
VAR_INPUT
    addRecipe    : BOOL;
    deleteRecipe : BOOL;
    modifyRecipe : BOOL;
    queryRecipe  : BOOL;
    recipeIn     : ST_Recipe;
END_VAR

VAR_OUTPUT
    recipeAdded       : BOOL := FALSE;
    recipeDeleted     : BOOL := FALSE;
    recipeModified    : BOOL := FALSE;
    recipeQueryResult : ST_Recipe;
    error             : BOOL := FALSE;
    status            : WORD := 0;
END_VAR

VAR_IN_OUT
    recipe : ARRAY[1..10] OF ST_Recipe;
END_VAR

VAR
    trigAdd    : R_TRIG;
    trigDelete : R_TRIG;
    trigModify : R_TRIG;
    trigQuery  : R_TRIG;
    tmp_i      : INT;
    tmp_slot   : INT;
    tmp_found  : BOOL;
    tmp_empty  : BOOL;
END_VAR

// Clear output flags at start of each scan
recipeAdded    := FALSE;
recipeDeleted  := FALSE;
recipeModified := FALSE;
error          := FALSE;
status         := 0;

// Detect rising edges on command inputs
trigQuery(CLK:=queryRecipe);
trigAdd(CLK:=addRecipe);
trigDelete(CLK:=deleteRecipe);
trigModify(CLK:=modifyRecipe);

// Operation 1: Query Recipe (PUB002, PUB008)
IF trigQuery.Q THEN
    tmp_found := FALSE;
    tmp_i := 1;
    WHILE tmp_i <= 10 AND NOT tmp_found DO
        IF recipe[tmp_i].recipeID = recipeIn.recipeID THEN
            tmp_found := TRUE;
        ELSE
            tmp_i := tmp_i + 1;
        END_IF;
    END_WHILE;

    IF tmp_found THEN
        recipeQueryResult := recipe[tmp_i];
        error   := FALSE;
        status  := 0;
    ELSE
        error   := TRUE;
        status  := 16#8001;  // Recipe not found
    END_IF;
END_IF;

// Operation 2: Add Recipe (PUB003, PUB009)
IF trigAdd.Q THEN
    // Check for duplicate recipeID
    tmp_found := FALSE;
    tmp_i := 1;
    WHILE tmp_i <= 10 AND NOT tmp_found DO
        IF recipe[tmp_i].recipeID = recipeIn.recipeID THEN
            tmp_found := TRUE;
        ELSE
            tmp_i := tmp_i + 1;
        END_IF;
    END_WHILE;

    IF tmp_found THEN
        error   := TRUE;
        status  := 16#8002;  // Duplicate recipeID
    ELSE
        // Find first empty slot (smallest index)
        tmp_empty := FALSE;
        tmp_slot  := 1;
        WHILE tmp_slot <= 10 AND NOT tmp_empty DO
            IF recipe[tmp_slot].recipeID = 0 THEN
                tmp_empty := TRUE;
            ELSE
                tmp_slot := tmp_slot + 1;
            END_IF;
        END_WHILE;

        IF tmp_empty THEN
            recipe[tmp_slot] := recipeIn;
            recipeAdded := TRUE;
            error       := FALSE;
            status      := 0;
        ELSE
            error   := TRUE;
            status  := 16#8003;  // No empty slot
        END_IF;
    END_IF;
END_IF;

// Operation 3: Delete Recipe (PUB004, PUB010)
IF trigDelete.Q THEN
    tmp_found := FALSE;
    tmp_i := 1;
    WHILE tmp_i <= 10 AND NOT tmp_found DO
        IF recipe[tmp_i].recipeID = recipeIn.recipeID THEN
            tmp_found := TRUE;
        ELSE
            tmp_i := tmp_i + 1;
        END_IF;
    END_WHILE;

    IF tmp_found THEN
        recipe[tmp_i].recipeID         := 0;
        recipe[tmp_i].ingredientType   := 0;
        recipe[tmp_i].ingredientRatio  := 0.0;
        recipe[tmp_i].productionTemperature := 0.0;
        recipeDeleted := TRUE;
        error         := FALSE;
        status        := 0;
    ELSE
        error   := TRUE;
        status  := 16#8004;  // Recipe not found for deletion
    END_IF;
END_IF;

// Operation 4: Modify Recipe (PUB005, PUB011)
IF trigModify.Q THEN
    tmp_found := FALSE;
    tmp_i := 1;
    WHILE tmp_i <= 10 AND NOT tmp_found DO
        IF recipe[tmp_i].recipeID = recipeIn.recipeID THEN
            tmp_found := TRUE;
        ELSE
            tmp_i := tmp_i + 1;
        END_IF;
    END_WHILE;

    IF tmp_found THEN
        recipe[tmp_i] := recipeIn;
        recipeModified := TRUE;
        error          := FALSE;
        status         := 0;
    ELSE
        error   := TRUE;
        status  := 16#8005;  // Recipe not found for modification
    END_IF;
END_IF;

END_FUNCTION_BLOCK

(* ---- public-hard-03.raw_candidate_01.st ---- *)
(* ENGINEERING_CONTRACT *)
(*
  Operation Priority (PUB001): Sequential evaluation order
    1. QUERY   - Read-only, sets recipeQueryResult
    2. ADD     - Write to empty slot, sets recipeAdded
    3. DELETE  - Write-clear slot, sets recipeDeleted
    4. MODIFY  - Write-replace slot, sets recipeModified

  Activation  : Edge-triggered via R_TRIG on command inputs
  Retention   : All outputs (except recipeQueryResult) are single-scan pulses
  Reset       : Outputs clear on subsequent scans when command deasserted
  Same-scan   : Final command state determines which R_TRIG fires
  Error       : error=TRUE with status code, no data written
  Success     : Specific success flag TRUE, error=FALSE, status=0
*)

(* CONTRACT_RULES [] *)

FUNCTION_BLOCK RecipeManagement
VAR_INPUT
    addRecipe    : BOOL;
    deleteRecipe : BOOL;
    modifyRecipe : BOOL;
    queryRecipe  : BOOL;
    recipeIn     : ST_Recipe;
END_VAR

VAR_OUTPUT
    recipeAdded       : BOOL := FALSE;
    recipeDeleted     : BOOL := FALSE;
    recipeModified    : BOOL := FALSE;
    recipeQueryResult : ST_Recipe;
    error             : BOOL := FALSE;
    status            : WORD := 0;
END_VAR

VAR_IN_OUT
    recipe : ARRAY[1..10] OF ST_Recipe;
END_VAR

VAR
    trigAdd    : R_TRIG;
    trigDelete : R_TRIG;
    trigModify : R_TRIG;
    trigQuery  : R_TRIG;
    tmp_i      : INT;
    tmp_slot   : INT;
    tmp_found  : BOOL;
    tmp_empty  : BOOL;
END_VAR

// Clear output flags at start of each scan
recipeAdded    := FALSE;
recipeDeleted  := FALSE;
recipeModified := FALSE;
error          := FALSE;
status         := 0;

// Detect rising edges on command inputs
trigQuery(IN:=queryRecipe);
trigAdd(IN:=addRecipe);
trigDelete(IN:=deleteRecipe);
trigModify(IN:=modifyRecipe);

// Operation 1: Query Recipe (PUB002, PUB008)
IF trigQuery.Q THEN
    tmp_found := FALSE;
    tmp_i := 1;
    WHILE tmp_i <= 10 AND NOT tmp_found DO
        IF recipe[tmp_i].recipeID = recipeIn.recipeID THEN
            tmp_found := TRUE;
        ELSE
            tmp_i := tmp_i + 1;
        END_IF;
    END_WHILE;

    IF tmp_found THEN
        recipeQueryResult := recipe[tmp_i];
        error   := FALSE;
        status  := 0;
    ELSE
        error   := TRUE;
        status  := 16#8001;  // Recipe not found
    END_IF;
END_IF;

// Operation 2: Add Recipe (PUB003, PUB009)
IF trigAdd.Q THEN
    // Check for duplicate recipeID
    tmp_found := FALSE;
    tmp_i := 1;
    WHILE tmp_i <= 10 AND NOT tmp_found DO
        IF recipe[tmp_i].recipeID = recipeIn.recipeID THEN
            tmp_found := TRUE;
        ELSE
            tmp_i := tmp_i + 1;
        END_IF;
    END_WHILE;

    IF tmp_found THEN
        error   := TRUE;
        status  := 16#8002;  // Duplicate recipeID
    ELSE
        // Find first empty slot (smallest index)
        tmp_empty := FALSE;
        tmp_slot  := 1;
        WHILE tmp_slot <= 10 AND NOT tmp_empty DO
            IF recipe[tmp_slot].recipeID = 0 THEN
                tmp_empty := TRUE;
            ELSE
                tmp_slot := tmp_slot + 1;
            END_IF;
        END_WHILE;

        IF tmp_empty THEN
            recipe[tmp_slot] := recipeIn;
            recipeAdded := TRUE;
            error       := FALSE;
            status      := 0;
        ELSE
            error   := TRUE;
            status  := 16#8003;  // No empty slot
        END_IF;
    END_IF;
END_IF;

// Operation 3: Delete Recipe (PUB004, PUB010)
IF trigDelete.Q THEN
    tmp_found := FALSE;
    tmp_i := 1;
    WHILE tmp_i <= 10 AND NOT tmp_found DO
        IF recipe[tmp_i].recipeID = recipeIn.recipeID THEN
            tmp_found := TRUE;
        ELSE
            tmp_i := tmp_i + 1;
        END_IF;
    END_WHILE;

    IF tmp_found THEN
        recipe[tmp_i].recipeID         := 0;
        recipe[tmp_i].ingredientType   := 0;
        recipe[tmp_i].ingredientRatio  := 0.0;
        recipe[tmp_i].productionTemperature := 0.0;
        recipeDeleted := TRUE;
        error         := FALSE;
        status        := 0;
    ELSE
        error   := TRUE;
        status  := 16#8004;  // Recipe not found for deletion
    END_IF;
END_IF;

// Operation 4: Modify Recipe (PUB005, PUB011)
IF trigModify.Q THEN
    tmp_found := FALSE;
    tmp_i := 1;
    WHILE tmp_i <= 10 AND NOT tmp_found DO
        IF recipe[tmp_i].recipeID = recipeIn.recipeID THEN
            tmp_found := TRUE;
        ELSE
            tmp_i := tmp_i + 1;
        END_IF;
    END_WHILE;

    IF tmp_found THEN
        recipe[tmp_i] := recipeIn;
        recipeModified := TRUE;
        error          := FALSE;
        status         := 0;
    ELSE
        error   := TRUE;
        status  := 16#8005;  // Recipe not found for modification
    END_IF;
END_IF;

END_FUNCTION_BLOCK

(* ---- public-hard-03.raw_candidate_02.st ---- *)
(* ENGINEERING_CONTRACT *)
(*
  Operation Priority (PUB001): Sequential evaluation order
    1. QUERY   - Read-only, sets recipeQueryResult
    2. ADD     - Write to empty slot, sets recipeAdded
    3. DELETE  - Write-clear slot, sets recipeDeleted
    4. MODIFY  - Write-replace slot, sets recipeModified

  Activation  : Edge-triggered via R_TRIG on command inputs
  Retention   : All outputs (except recipeQueryResult) are single-scan pulses
  Reset       : Outputs clear on subsequent scans when command deasserted
  Same-scan   : Final command state determines which R_TRIG fires
  Error       : error=TRUE with status code, no data written
  Success     : Specific success flag TRUE, error=FALSE, status=0
*)

TYPE ST_Recipe : STRUCT
    recipeID              : INT;
    ingredientType        : INT;
    ingredientRatio       : REAL;
    productionTemperature : REAL;
END_STRUCT END_TYPE

(* CONTRACT_RULES [] *)

FUNCTION_BLOCK RecipeManagement
VAR_INPUT
    addRecipe    : BOOL;
    deleteRecipe : BOOL;
    modifyRecipe : BOOL;
    queryRecipe  : BOOL;
    recipeIn     : ST_Recipe;
END_VAR

VAR_OUTPUT
    recipeAdded       : BOOL := FALSE;
    recipeDeleted     : BOOL := FALSE;
    recipeModified    : BOOL := FALSE;
    recipeQueryResult : ST_Recipe;
    error             : BOOL := FALSE;
    status            : WORD := 0;
END_VAR

VAR_IN_OUT
    recipe : ARRAY[1..10] OF ST_Recipe;
END_VAR

VAR
    trigAdd    : R_TRIG;
    trigDelete : R_TRIG;
    trigModify : R_TRIG;
    trigQuery  : R_TRIG;
    tmp_i      : INT;
    tmp_slot   : INT;
    tmp_found  : BOOL;
    tmp_empty  : BOOL;
END_VAR

// Clear output flags at start of each scan
recipeAdded    := FALSE;
recipeDeleted  := FALSE;
recipeModified := FALSE;
error          := FALSE;
status         := 0;

// Detect rising edges on command inputs
trigQuery(CLK:=queryRecipe);
trigAdd(CLK:=addRecipe);
trigDelete(CLK:=deleteRecipe);
trigModify(CLK:=modifyRecipe);

// Operation 1: Query Recipe (PUB002, PUB008)
IF trigQuery.Q THEN
    tmp_found := FALSE;
    tmp_i := 1;
    WHILE tmp_i <= 10 AND NOT tmp_found DO
        IF recipe[tmp_i].recipeID = recipeIn.recipeID THEN
            tmp_found := TRUE;
        ELSE
            tmp_i := tmp_i + 1;
        END_IF;
    END_WHILE;

    IF tmp_found THEN
        recipeQueryResult := recipe[tmp_i];
        error   := FALSE;
        status  := 0;
    ELSE
        error   := TRUE;
        status  := 16#8001;  // Recipe not found
    END_IF;
END_IF;

// Operation 2: Add Recipe (PUB003, PUB009)
IF trigAdd.Q THEN
    // Check for duplicate recipeID
    tmp_found := FALSE;
    tmp_i := 1;
    WHILE tmp_i <= 10 AND NOT tmp_found DO
        IF recipe[tmp_i].recipeID = recipeIn.recipeID THEN
            tmp_found := TRUE;
        ELSE
            tmp_i := tmp_i + 1;
        END_IF;
    END_WHILE;

    IF tmp_found THEN
        error   := TRUE;
        status  := 16#8002;  // Duplicate recipeID
    ELSE
        // Find first empty slot (smallest index)
        tmp_empty := FALSE;
        tmp_slot  := 1;
        WHILE tmp_slot <= 10 AND NOT tmp_empty DO
            IF recipe[tmp_slot].recipeID = 0 THEN
                tmp_empty := TRUE;
            ELSE
                tmp_slot := tmp_slot + 1;
            END_IF;
        END_WHILE;

        IF tmp_empty THEN
            recipe[tmp_slot] := recipeIn;
            recipeAdded := TRUE;
            error       := FALSE;
            status      := 0;
        ELSE
            error   := TRUE;
            status  := 16#8003;  // No empty slot
        END_IF;
    END_IF;
END_IF;

// Operation 3: Delete Recipe (PUB004, PUB010)
IF trigDelete.Q THEN
    tmp_found := FALSE;
    tmp_i := 1;
    WHILE tmp_i <= 10 AND NOT tmp_found DO
        IF recipe[tmp_i].recipeID = recipeIn.recipeID THEN
            tmp_found := TRUE;
        ELSE
            tmp_i := tmp_i + 1;
        END_IF;
    END_WHILE;

    IF tmp_found THEN
        recipe[tmp_i].recipeID         := 0;
        recipe[tmp_i].ingredientType   := 0;
        recipe[tmp_i].ingredientRatio  := 0.0;
        recipe[tmp_i].productionTemperature := 0.0;
        recipeDeleted := TRUE;
        error         := FALSE;
        status        := 0;
    ELSE
        error   := TRUE;
        status  := 16#8004;  // Recipe not found for deletion
    END_IF;
END_IF;

// Operation 4: Modify Recipe (PUB005, PUB011)
IF trigModify.Q THEN
    tmp_found := FALSE;
    tmp_i := 1;
    WHILE tmp_i <= 10 AND NOT tmp_found DO
        IF recipe[tmp_i].recipeID = recipeIn.recipeID THEN
            tmp_found := TRUE;
        ELSE
            tmp_i := tmp_i + 1;
        END_IF;
    END_WHILE;

    IF tmp_found THEN
        recipe[tmp_i] := recipeIn;
        recipeModified := TRUE;
        error          := FALSE;
        status         := 0;
    ELSE
        error   := TRUE;
        status  := 16#8005;  // Recipe not found for modification
    END_IF;
END_IF;

END_FUNCTION_BLOCK

(* ---- public-hard-03.raw_candidate_04.st ---- *)
(* ENGINEERING_CONTRACT *)
(*
  Operation Priority (PUB001): Sequential evaluation order
    1. QUERY   - Read-only, sets recipeQueryResult
    2. ADD     - Write to empty slot, sets recipeAdded
    3. DELETE  - Write-clear slot, sets recipeDeleted
    4. MODIFY  - Write-replace slot, sets recipeModified

  Activation  : Edge-triggered via R_TRIG on command inputs
  Retention   : All outputs (except recipeQueryResult) are single-scan pulses
  Reset       : Outputs clear on subsequent scans when command deasserted
  Same-scan   : Final command state determines which R_TRIG fires
  Error       : error=TRUE with status code, no data written
  Success     : Specific success flag TRUE, error=FALSE, status=0
*)

TYPE ST_Recipe : STRUCT
    recipeID              : INT;
    ingredientType        : INT;
    ingredientRatio       : REAL;
    productionTemperature : REAL;
END_STRUCT END_TYPE;

(* CONTRACT_RULES [] *)

FUNCTION_BLOCK RecipeManagement
VAR_INPUT
    addRecipe    : BOOL;
    deleteRecipe : BOOL;
    modifyRecipe : BOOL;
    queryRecipe  : BOOL;
    recipeIn     : ST_Recipe;
END_VAR

VAR_OUTPUT
    recipeAdded       : BOOL := FALSE;
    recipeDeleted     : BOOL := FALSE;
    recipeModified    : BOOL := FALSE;
    recipeQueryResult : ST_Recipe;
    error             : BOOL := FALSE;
    status            : WORD := 0;
END_VAR

VAR_IN_OUT
    recipe : ARRAY[1..10] OF ST_Recipe;
END_VAR

VAR
    trigAdd    : R_TRIG;
    trigDelete : R_TRIG;
    trigModify : R_TRIG;
    trigQuery  : R_TRIG;
    tmp_i      : INT;
    tmp_slot   : INT;
    tmp_found  : BOOL;
    tmp_empty  : BOOL;
END_VAR

// Clear output flags at start of each scan
recipeAdded    := FALSE;
recipeDeleted  := FALSE;
recipeModified := FALSE;
IF trigQuery.Q OR trigAdd.Q OR trigDelete.Q OR trigModify.Q THEN
    error   := FALSE;
    status  := 0;
END_IF;

// Detect rising edges on command inputs
trigQuery(CLK:=queryRecipe);
trigAdd(CLK:=addRecipe);
trigDelete(CLK:=deleteRecipe);
trigModify(CLK:=modifyRecipe);

// Operation 1: Query Recipe (PUB002, PUB008)
IF trigQuery.Q THEN
    tmp_found := FALSE;
    tmp_i := 1;
    WHILE tmp_i <= 10 AND NOT tmp_found DO
        IF recipe[tmp_i].recipeID = recipeIn.recipeID THEN
            tmp_found := TRUE;
        ELSE
            tmp_i := tmp_i + 1;
        END_IF;
    END_WHILE;

    IF tmp_found THEN
        recipeQueryResult := recipe[tmp_i];
        error   := FALSE;
        status  := 0;
    ELSE
        error   := TRUE;
        status  := 16#8001;  // Recipe not found
    END_IF;
END_IF;

// Operation 2: Add Recipe (PUB003, PUB009)
IF trigAdd.Q THEN
    // Check for duplicate recipeID
    tmp_found := FALSE;
    tmp_i := 1;
    WHILE tmp_i <= 10 AND NOT tmp_found DO
        IF recipe[tmp_i].recipeID = recipeIn.recipeID THEN
            tmp_found := TRUE;
        ELSE
            tmp_i := tmp_i + 1;
        END_IF;
    END_WHILE;

    IF tmp_found THEN
        error   := TRUE;
        status  := 16#8002;  // Duplicate recipeID
    ELSE
        // Find first empty slot (smallest index)
        tmp_empty := FALSE;
        tmp_slot  := 1;
        WHILE tmp_slot <= 10 AND NOT tmp_empty DO
            IF recipe[tmp_slot].recipeID = 0 THEN
                tmp_empty := TRUE;
            ELSE
                tmp_slot := tmp_slot + 1;
            END_IF;
        END_WHILE;

        IF tmp_empty THEN
            recipe[tmp_slot] := recipeIn;
            recipeAdded := TRUE;
            error       := FALSE;
            status      := 0;
        ELSE
            error   := TRUE;
            status  := 16#8003;  // No empty slot
        END_IF;
    END_IF;
END_IF;

// Operation 3: Delete Recipe (PUB004, PUB010)
IF trigDelete.Q THEN
    tmp_found := FALSE;
    tmp_i := 1;
    WHILE tmp_i <= 10 AND NOT tmp_found DO
        IF recipe[tmp_i].recipeID = recipeIn.recipeID THEN
            tmp_found := TRUE;
        ELSE
            tmp_i := tmp_i + 1;
        END_IF;
    END_WHILE;

    IF tmp_found THEN
        recipe[tmp_i].recipeID         := 0;
        recipe[tmp_i].ingredientType   := 0;
        recipe[tmp_i].ingredientRatio  := 0.0;
        recipe[tmp_i].productionTemperature := 0.0;
        recipeDeleted := TRUE;
        error         := FALSE;
        status        := 0;
    ELSE
        error   := TRUE;
        status  := 16#8004;  // Recipe not found for deletion
    END_IF;
END_IF;

// Operation 4: Modify Recipe (PUB005, PUB011)
IF trigModify.Q THEN
    tmp_found := FALSE;
    tmp_i := 1;
    WHILE tmp_i <= 10 AND NOT tmp_found DO
        IF recipe[tmp_i].recipeID = recipeIn.recipeID THEN
            tmp_found := TRUE;
        ELSE
            tmp_i := tmp_i + 1;
        END_IF;
    END_WHILE;

    IF tmp_found THEN
        recipe[tmp_i] := recipeIn;
        recipeModified := TRUE;
        error          := FALSE;
        status         := 0;
    ELSE
        error   := TRUE;
        status  := 16#8005;  // Recipe not found for modification
    END_IF;
END_IF;

END_FUNCTION_BLOCK

(* ---- public-hard-04.candidate_01.st ---- *)
// FIFO Queue Implementation - CODESYS 3.5
// PUB001: Rising edge enqueue appends item to tail if not full
// PUB002: Rising edge dequeue removes front to item if not empty; caller must not combine enq+deq
// PUB003: reset=TRUE empties queue, sets elementCount=0; takes priority; buffer values may persist
// PUB004: elementCount=0..capacity; 0=empty, capacity=full
// PUB005: Reject deq when empty or enq when full; leave queue/item unchanged; status reports reason
// PUB006: status=16#0000(no err), 16#8001(deq rejected empty), 16#8002(enq rejected full)
// Internal: First invocation derives capacity; circular queue with head/tail; R_TRIG for edges

FUNCTION_BLOCK FB_FIFOQueue
VAR_INPUT
    enqueue  : BOOL;
    dequeue  : BOOL;
    reset    : BOOL;
END_VAR

VAR_OUTPUT
    elementCount : DINT := 0;
    status       : WORD := 16#0000;
END_VAR

VAR_IN_OUT
    item   : VARIANT;
    buffer : VARIANT;
END_VAR

VAR
    R_Trig_Reset   : R_TRIG;
    R_Trig_Enqueue : R_TRIG;
    R_Trig_Dequeue : R_TRIG;
    head           : DINT := 0;
    tail           : DINT := 0;
    count          : DINT := 0;
    capacity       : DINT := 0;
    tmp_Item       : DINT;
    tmp_Index      : DINT;
    tmp_FirstScan  : BOOL := TRUE;
END_VAR

(* CONTRACT_RULES [] *)

IF tmp_FirstScan THEN
    tmp_FirstScan := FALSE;
    tmp_Index := UPPER_BOUND(buffer, 1) - LOWER_BOUND(buffer, 1);
    capacity := DINT_TO_INT(tmp_Index) + 1;
    head := 0;
    tail := 0;
    count := 0;
END_IF;

R_Trig_Reset(CLK := reset);
R_Trig_Enqueue(CLK := enqueue);
R_Trig_Dequeue(CLK := dequeue);

IF R_Trig_Reset.Q THEN
    count := 0;
    head := 0;
    tail := 0;
    elementCount := 0;
    status := 16#0000;
    RETURN;
END_IF;

IF R_Trig_Enqueue.Q THEN
    IF count >= capacity THEN
        status := 16#8002;
        RETURN;
    END_IF;
    tmp_Item := VARIANT_TO_DINT(item);
    tmp_Index := LOWER_BOUND(buffer, 1) + tail;
    buffer[tmp_Index] := DINT_TO_VARIANT(tmp_Item);
    tail := (tail + 1) MOD capacity;
    count := count + 1;
    elementCount := count;
    status := 16#0000;
    RETURN;
END_IF;

IF R_Trig_Dequeue.Q THEN
    IF count <= 0 THEN
        status := 16#8001;
        RETURN;
    END_IF;
    tmp_Index := LOWER_BOUND(buffer, 1) + head;
    tmp_Item := VARIANT_TO_DINT(buffer[tmp_Index]);
    item := DINT_TO_VARIANT(tmp_Item);
    head := (head + 1) MOD capacity;
    count := count - 1;
    elementCount := count;
    status := 16#0000;
    RETURN;
END_IF;

elementCount := count;
status := 16#0000;

END_FUNCTION_BLOCK

(* ---- public-hard-04.raw_candidate_01.st ---- *)
// FIFO Queue Implementation - CODESYS 3.5
// PUB001: Rising edge enqueue appends item to tail if not full
// PUB002: Rising edge dequeue removes front to item if not empty; caller must not combine enq+deq
// PUB003: reset=TRUE empties queue, sets elementCount=0; takes priority; buffer values may persist
// PUB004: elementCount=0..capacity; 0=empty, capacity=full
// PUB005: Reject deq when empty or enq when full; leave queue/item unchanged; status reports reason
// PUB006: status=16#0000(no err), 16#8001(deq rejected empty), 16#8002(enq rejected full)
// Internal: First invocation derives capacity; circular queue with head/tail; R_TRIG for edges

FUNCTION_BLOCK FB_FIFOQueue
VAR_INPUT
    enqueue  : BOOL;
    dequeue  : BOOL;
    reset    : BOOL;
END_VAR

VAR_OUTPUT
    elementCount : DINT := 0;
    status       : WORD := 16#0000;
END_VAR

VAR_IN_OUT
    item   : VARIANT;
    buffer : VARIANT;
END_VAR

VAR
    R_Trig_Reset   : R_TRIG;
    R_Trig_Enqueue : R_TRIG;
    R_Trig_Dequeue : R_TRIG;
    head           : DINT := 0;
    tail           : DINT := 0;
    count          : DINT := 0;
    capacity       : DINT := 0;
    tmp_Item       : DINT;
    tmp_Index      : DINT;
    tmp_FirstScan  : BOOL := TRUE;
END_VAR

(* CONTRACT_RULES [] *)

IF tmp_FirstScan THEN
    tmp_FirstScan := FALSE;
    tmp_Index := UPPER_BOUND(buffer, 1) - LOWER_BOUND(buffer, 1);
    capacity := DINT_TO_INT(tmp_Index) + 1;
    head := 0;
    tail := 0;
    count := 0;
END_IF

R_Trig_Reset(CLK := reset);
R_Trig_Enqueue(CLK := enqueue);
R_Trig_Dequeue(CLK := dequeue);

IF R_Trig_Reset.Q THEN
    count := 0;
    head := 0;
    tail := 0;
    elementCount := 0;
    status := 16#0000;
    RETURN;
END_IF

IF R_Trig_Enqueue.Q THEN
    IF count >= capacity THEN
        status := 16#8002;
        RETURN;
    END_IF
    tmp_Item := VARIANT_TO_DINT(item);
    tmp_Index := LOWER_BOUND(buffer, 1) + tail;
    buffer[tmp_Index] := DINT_TO_VARIANT(tmp_Item);
    tail := (tail + 1) MOD capacity;
    count := count + 1;
    elementCount := count;
    status := 16#0000;
    RETURN;
END_IF

IF R_Trig_Dequeue.Q THEN
    IF count <= 0 THEN
        status := 16#8001;
        RETURN;
    END_IF
    tmp_Index := LOWER_BOUND(buffer, 1) + head;
    tmp_Item := VARIANT_TO_DINT(buffer[tmp_Index]);
    item := DINT_TO_VARIANT(tmp_Item);
    head := (head + 1) MOD capacity;
    count := count - 1;
    elementCount := count;
    status := 16#0000;
    RETURN;
END_IF

elementCount := count;
status := 16#0000;

END_FUNCTION_BLOCK

(* ---- public-hard-05.candidate_01.st ---- *)
(* ENGINEERING_CONTRACT *)
(*
  PUB001: Manual mode - button activates output while held, stop at limit switch or release.
          Manual outputs: retention=hold_until_button_release OR limit, reset=button_release OR limit_reached.
  PUB002: Emergency stop - all outputs OFF, all state cleared. No retention. Reset=EmergencyStop=TRUE.
  PUB003-PUB012: Single step mode - 8-step sequence, Start to advance each step.
          Step outputs: retention=hold_until_limit, reset=limit_reached OR mode_exit.
          Step index 1..8 maps to: Down→Grip→Up→Right→Down→Release→Up→Left→(repeat).
  PUB013-PUB014: Single cycle mode - auto-execute 8 steps on Start, stop at home.
          Same output retention as PUB003-PUB012. Cycle reset=mode_exit only.
  PUB015-PUB016: Continuous mode - same as single cycle but repeat after home.
          Cycle restart trigger: timer PT after home, if Start still asserted.
  PUB017: GripLimitSwitch/ReleaseLimitSwitch signal action completion (not position).
          Grip/Release output: activation=entry_unless_limit, retention=limit FALSE,
          deactivation=limit TRUE (same scan). No explicit reset input.
  PUB018: Caller guarantees mutually exclusive mode inputs.
  PUB019: Opposite-direction pairs (Up/Down, Left/Right) must never energize together.
          Implementation: output TRUE only when opposite limit is FALSE.
  PUB020: Single step confirmation = Start button release, not level.
*)
(* CONTRACT_RULES [] *)

TYPE ArmStep : INT (Idle := 0, Step1 := 1, Step2 := 2, Step3 := 3, Step4 := 4,
                     Step5 := 5, Step6 := 6, Step7 := 7, Step8 := 8)
END_TYPE;

FUNCTION_BLOCK ArmController
VAR_INPUT
    ManualMode       : BOOL;
    SingleStepMode   : BOOL;
    SingleCycleMode  : BOOL;
    ContinuousMode   : BOOL;
    EmergencyStop    : BOOL;
    Start            : BOOL;
    DownButton       : BOOL;
    UpButton         : BOOL;
    LeftButton       : BOOL;
    RightButton      : BOOL;
    GripButton       : BOOL;
    ReleaseButton    : BOOL;
    DownLimitSwitch  : BOOL;
    UpLimitSwitch    : BOOL;
    LeftLimitSwitch  : BOOL;
    RightLimitSwitch : BOOL;
    GripLimitSwitch  : BOOL;
    ReleaseLimitSwitch : BOOL;
END_VAR
VAR_OUTPUT
    MoveDown       : BOOL;
    MoveUp         : BOOL;
    MoveLeft       : BOOL;
    MoveRight      : BOOL;
    ActivateGrip   : BOOL;
    ActivateRelease : BOOL;
END_VAR
VAR
    tmp_CurrentStep   : ArmStep := ArmStep.Idle;
    tmp_StartTrigger  : BOOL;
    tmp_StartReleased : BOOL;
    tmp_Gripping      : BOOL;
    tmp_Releasing     : BOOL;
    tmp_CycleDoneTimer : TON;
END_VAR

// Emergency stop: clears all outputs and state
IF EmergencyStop THEN
    MoveDown       := FALSE;
    MoveUp         := FALSE;
    MoveLeft       := FALSE;
    MoveRight      := FALSE;
    ActivateGrip   := FALSE;
    ActivateRelease := FALSE;
    tmp_CurrentStep   := ArmStep.Idle;
    tmp_StartTrigger  := FALSE;
    tmp_StartReleased := FALSE;
    tmp_Gripping      := FALSE;
    tmp_Releasing     := FALSE;
    tmp_CycleDoneTimer(IN := FALSE, PT := T#0s);
    RETURN;
END_IF;

// Default all outputs OFF
MoveDown       := FALSE;
MoveUp         := FALSE;
MoveLeft       := FALSE;
MoveRight      := FALSE;
ActivateGrip   := FALSE;
ActivateRelease := FALSE;

IF ManualMode THEN
    // Direct button-to-output mapping, stop at limit switch
    MoveDown       := DownButton AND NOT DownLimitSwitch;
    MoveUp         := UpButton AND NOT UpLimitSwitch;
    MoveLeft       := LeftButton AND NOT LeftLimitSwitch;
    MoveRight      := RightButton AND NOT RightLimitSwitch;
    ActivateGrip   := GripButton AND NOT GripLimitSwitch;
    ActivateRelease := ReleaseButton AND NOT ReleaseLimitSwitch;

ELSIF SingleStepMode THEN
    // Rising-edge Start advances through steps; each step waits for limit switch
    IF tmp_StartReleased AND NOT Start AND tmp_CurrentStep = ArmStep.Idle THEN
        tmp_StartTrigger := TRUE;
    END_IF;
    tmp_StartReleased := Start;

    IF tmp_CurrentStep = ArmStep.Idle THEN
        IF tmp_StartTrigger THEN
            tmp_CurrentStep := ArmStep.Step1;
            tmp_StartTrigger := FALSE;
        END_IF;
    ELSE
        CASE TO_INT(tmp_CurrentStep) OF
            1: MoveDown := NOT DownLimitSwitch;
               IF DownLimitSwitch THEN
                   tmp_CurrentStep := ArmStep.Step2;
               END_IF;
            2: ActivateGrip := NOT GripLimitSwitch;
               IF GripLimitSwitch THEN
                   tmp_CurrentStep := ArmStep.Step3;
               END_IF;
            3: MoveUp := NOT UpLimitSwitch;
               IF UpLimitSwitch THEN
                   tmp_CurrentStep := ArmStep.Step4;
               END_IF;
            4: MoveRight := NOT RightLimitSwitch;
               IF RightLimitSwitch THEN
                   tmp_CurrentStep := ArmStep.Step5;
               END_IF;
            5: MoveDown := NOT DownLimitSwitch;
               IF DownLimitSwitch THEN
                   tmp_CurrentStep := ArmStep.Step6;
               END_IF;
            6: ActivateRelease := NOT ReleaseLimitSwitch;
               IF ReleaseLimitSwitch THEN
                   tmp_CurrentStep := ArmStep.Step7;
               END_IF;
            7: MoveUp := NOT UpLimitSwitch;
               IF UpLimitSwitch THEN
                   tmp_CurrentStep := ArmStep.Step8;
               END_IF;
            8: MoveLeft := NOT LeftLimitSwitch;
               IF LeftLimitSwitch THEN
                   tmp_CurrentStep := ArmStep.Idle;
               END_IF;
        END_CASE;
    END_IF;

ELSIF SingleCycleMode THEN
    // Start triggers auto-sequence; cycle completes and stops at home
    IF Start AND tmp_CurrentStep = ArmStep.Idle AND NOT tmp_Gripping AND NOT tmp_Releasing THEN
        tmp_StartTrigger := TRUE;
    END_IF;

    // Cycle completion: at Step8 and home (UpLimitSwitch AND LeftLimitSwitch)
    IF tmp_CurrentStep = ArmStep.Step8 AND UpLimitSwitch AND LeftLimitSwitch THEN
        tmp_CycleDoneTimer(IN := TRUE, PT := T#1ms);
        IF tmp_CycleDoneTimer.Q THEN
            tmp_StartTrigger  := FALSE;
            tmp_Gripping      := FALSE;
            tmp_Releasing     := FALSE;
            tmp_CurrentStep   := ArmStep.Idle;
        END_IF;
    ELSE
        tmp_CycleDoneTimer(IN := FALSE, PT := T#0s);
    END_IF;

    IF tmp_StartTrigger THEN
        CASE TO_INT(tmp_CurrentStep) OF
            0: tmp_CurrentStep := ArmStep.Step1;
            1: MoveDown := NOT DownLimitSwitch;
               IF DownLimitSwitch THEN
                   tmp_CurrentStep := ArmStep.Step2;
               END_IF;
            2: ActivateGrip := NOT GripLimitSwitch;
               IF GripLimitSwitch THEN
                   tmp_CurrentStep := ArmStep.Step3;
               END_IF;
            3: MoveUp := NOT UpLimitSwitch;
               IF UpLimitSwitch THEN
                   tmp_CurrentStep := ArmStep.Step4;
               END_IF;
            4: MoveRight := NOT RightLimitSwitch;
               IF RightLimitSwitch THEN
                   tmp_CurrentStep := ArmStep.Step5;
               END_IF;
            5: MoveDown := NOT DownLimitSwitch;
               IF DownLimitSwitch THEN
                   tmp_CurrentStep := ArmStep.Step6;
               END_IF;
            6: ActivateRelease := NOT ReleaseLimitSwitch;
               IF ReleaseLimitSwitch THEN
                   tmp_CurrentStep := ArmStep.Step7;
               END_IF;
            7: MoveUp := NOT UpLimitSwitch;
               IF UpLimitSwitch THEN
                   tmp_CurrentStep := ArmStep.Step8;
               END_IF;
            8: MoveLeft := NOT LeftLimitSwitch;
               IF LeftLimitSwitch THEN
                   tmp_CurrentStep := ArmStep.Idle;
               END_IF;
        END_CASE;
    END_IF;

ELSIF ContinuousMode THEN
    // Same as single cycle but restarts automatically after PT delay at home
    IF Start AND NOT tmp_Gripping AND NOT tmp_Releasing THEN
        tmp_StartTrigger := TRUE;
    END_IF;

    IF tmp_CurrentStep = ArmStep.Step8 AND UpLimitSwitch AND LeftLimitSwitch THEN
        tmp_CycleDoneTimer(IN := tmp_CycleDoneTimer.Q, PT := T#1ms);
        IF tmp_CycleDoneTimer.Q THEN
            tmp_CurrentStep := ArmStep.Idle;
        END_IF;
        IF NOT tmp_CycleDoneTimer.Q AND tmp_CurrentStep = ArmStep.Idle THEN
            tmp_StartTrigger := Start;
            tmp_Gripping     := FALSE;
            tmp_Releasing    := FALSE;
        END_IF;
    ELSE
        tmp_CycleDoneTimer(IN := FALSE, PT := T#0s);
    END_IF;

    IF tmp_StartTrigger THEN
        CASE TO_INT(tmp_CurrentStep) OF
            0: tmp_CurrentStep := ArmStep.Step1;
            1: MoveDown := NOT DownLimitSwitch;
               IF DownLimitSwitch THEN
                   tmp_CurrentStep := ArmStep.Step2;
               END_IF;
            2: ActivateGrip := NOT GripLimitSwitch;
               IF GripLimitSwitch THEN
                   tmp_CurrentStep := ArmStep.Step3;
               END_IF;
            3: MoveUp := NOT UpLimitSwitch;
               IF UpLimitSwitch THEN
                   tmp_CurrentStep := ArmStep.Step4;
               END_IF;
            4: MoveRight := NOT RightLimitSwitch;
               IF RightLimitSwitch THEN
                   tmp_CurrentStep := ArmStep.Step5;
               END_IF;
            5: MoveDown := NOT DownLimitSwitch;
               IF DownLimitSwitch THEN
                   tmp_CurrentStep := ArmStep.Step6;
               END_IF;
            6: ActivateRelease := NOT ReleaseLimitSwitch;
               IF ReleaseLimitSwitch THEN
                   tmp_CurrentStep := ArmStep.Step7;
               END_IF;
            7: MoveUp := NOT UpLimitSwitch;
               IF UpLimitSwitch THEN
                   tmp_CurrentStep := ArmStep.Step8;
               END_IF;
            8: MoveLeft := NOT LeftLimitSwitch;
               IF LeftLimitSwitch THEN
                   tmp_CurrentStep := ArmStep.Idle;
               END_IF;
        END_CASE;
    END_IF;
END_IF;

END_FUNCTION_BLOCK

(* ---- public-hard-05.patch_base_02.st ---- *)
(* ENGINEERING_CONTRACT *)
(*
  PUB001: Manual mode - button activates output while held, stop at limit switch or release.
          Manual outputs: retention=hold_until_button_release OR limit, reset=button_release OR limit_reached.
  PUB002: Emergency stop - all outputs OFF, all state cleared. No retention. Reset=EmergencyStop=TRUE.
  PUB003-PUB012: Single step mode - 8-step sequence, Start to advance each step.
          Step outputs: retention=hold_until_limit, reset=limit_reached OR mode_exit.
          Step index 1..8 maps to: Down→Grip→Up→Right→Down→Release→Up→Left→(repeat).
  PUB013-PUB014: Single cycle mode - auto-execute 8 steps on Start, stop at home.
          Same output retention as PUB003-PUB012. Cycle reset=mode_exit only.
  PUB015-PUB016: Continuous mode - same as single cycle but repeat after home.
          Cycle restart trigger: timer PT after home, if Start still asserted.
  PUB017: GripLimitSwitch/ReleaseLimitSwitch signal action completion (not position).
          Grip/Release output: activation=entry_unless_limit, retention=limit FALSE,
          deactivation=limit TRUE (same scan). No explicit reset input.
  PUB018: Caller guarantees mutually exclusive mode inputs.
  PUB019: Opposite-direction pairs (Up/Down, Left/Right) must never energize together.
          Implementation: output TRUE only when opposite limit is FALSE.
  PUB020: Single step confirmation = Start button release, not level.
*)
(* CONTRACT_RULES [] *)

TYPE ArmStep : INT (Idle := 0, Step1 := 1, Step2 := 2, Step3 := 3, Step4 := 4,
                     Step5 := 5, Step6 := 6, Step7 := 7, Step8 := 8)
END_TYPE;

FUNCTION_BLOCK ArmController
VAR_INPUT
    ManualMode       : BOOL;
    SingleStepMode   : BOOL;
    SingleCycleMode  : BOOL;
    ContinuousMode   : BOOL;
    EmergencyStop    : BOOL;
    Start            : BOOL;
    DownButton       : BOOL;
    UpButton         : BOOL;
    LeftButton       : BOOL;
    RightButton      : BOOL;
    GripButton       : BOOL;
    ReleaseButton    : BOOL;
    DownLimitSwitch  : BOOL;
    UpLimitSwitch    : BOOL;
    LeftLimitSwitch  : BOOL;
    RightLimitSwitch : BOOL;
    GripLimitSwitch  : BOOL;
    ReleaseLimitSwitch : BOOL;
END_VAR
VAR_OUTPUT
    MoveDown       : BOOL;
    MoveUp         : BOOL;
    MoveLeft       : BOOL;
    MoveRight      : BOOL;
    ActivateGrip   : BOOL;
    ActivateRelease : BOOL;
END_VAR
VAR
    tmp_CurrentStep   : ArmStep := ArmStep.Idle;
    tmp_StartTrigger  : BOOL;
    tmp_StartReleased : BOOL;
    tmp_Gripping      : BOOL;
    tmp_Releasing     : BOOL;
    tmp_CycleDoneTimer : TON;
END_VAR

// Emergency stop: clears all outputs and state
IF EmergencyStop THEN
    MoveDown       := FALSE;
    MoveUp         := FALSE;
    MoveLeft       := FALSE;
    MoveRight      := FALSE;
    ActivateGrip   := FALSE;
    ActivateRelease := FALSE;
    tmp_CurrentStep   := ArmStep.Idle;
    tmp_StartTrigger  := FALSE;
    tmp_StartReleased := FALSE;
    tmp_Gripping      := FALSE;
    tmp_Releasing     := FALSE;
    tmp_CycleDoneTimer(IN := FALSE, PT := T#0s);
    RETURN;
END_IF;

// Default all outputs OFF
MoveDown       := FALSE;
MoveUp         := FALSE;
MoveLeft       := FALSE;
MoveRight      := FALSE;
ActivateGrip   := FALSE;
ActivateRelease := FALSE;

IF ManualMode THEN
    // Direct button-to-output mapping, stop at limit switch
    MoveDown       := DownButton AND NOT DownLimitSwitch;
    MoveUp         := UpButton AND NOT UpLimitSwitch;
    MoveLeft       := LeftButton AND NOT LeftLimitSwitch;
    MoveRight      := RightButton AND NOT RightLimitSwitch;
    ActivateGrip   := GripButton AND NOT GripLimitSwitch;
    ActivateRelease := ReleaseButton AND NOT ReleaseLimitSwitch;

ELSIF SingleStepMode THEN
    // Rising-edge Start advances through steps; each step waits for limit switch
    IF tmp_StartReleased AND NOT Start AND tmp_CurrentStep = ArmStep.Idle THEN
        tmp_StartTrigger := TRUE;
    END_IF;
    tmp_StartReleased := Start;

    IF tmp_CurrentStep = ArmStep.Idle THEN
        IF tmp_StartTrigger THEN
            tmp_CurrentStep := ArmStep.Step1;
            tmp_StartTrigger := FALSE;
        END_IF;
    ELSE
        CASE TO_INT(tmp_CurrentStep) OF
            1: MoveDown := NOT DownLimitSwitch;
               IF DownLimitSwitch THEN
                   tmp_CurrentStep := ArmStep.Step2;
               END_IF;
            2: ActivateGrip := NOT GripLimitSwitch;
               IF GripLimitSwitch THEN
                   tmp_CurrentStep := ArmStep.Step3;
               END_IF;
            3: MoveUp := NOT UpLimitSwitch;
               IF UpLimitSwitch THEN
                   tmp_CurrentStep := ArmStep.Step4;
               END_IF;
            4: MoveRight := NOT RightLimitSwitch;
               IF RightLimitSwitch THEN
                   tmp_CurrentStep := ArmStep.Step5;
               END_IF;
            5: MoveDown := NOT DownLimitSwitch;
               IF DownLimitSwitch THEN
                   tmp_CurrentStep := ArmStep.Step6;
               END_IF;
            6: ActivateRelease := NOT ReleaseLimitSwitch;
               IF ReleaseLimitSwitch THEN
                   tmp_CurrentStep := ArmStep.Step7;
               END_IF;
            7: MoveUp := NOT UpLimitSwitch;
               IF UpLimitSwitch THEN
                   tmp_CurrentStep := ArmStep.Step8;
               END_IF;
            8: MoveLeft := NOT LeftLimitSwitch;
               IF LeftLimitSwitch THEN
                   tmp_CurrentStep := ArmStep.Idle;
               END_IF;
        END_CASE;
    END_IF;

ELSIF SingleCycleMode THEN
    // Start triggers auto-sequence; cycle completes and stops at home
    IF Start AND tmp_CurrentStep = ArmStep.Idle AND NOT tmp_Gripping AND NOT tmp_Releasing THEN
        tmp_StartTrigger := TRUE;
    END_IF;

    // Cycle completion: at Step8 and home (UpLimitSwitch AND LeftLimitSwitch)
    IF tmp_CurrentStep = ArmStep.Step8 AND UpLimitSwitch AND LeftLimitSwitch THEN
        tmp_CycleDoneTimer(IN := TRUE, PT := T#1ms);
        IF tmp_CycleDoneTimer.Q THEN
            tmp_StartTrigger  := FALSE;
            tmp_Gripping      := FALSE;
            tmp_Releasing     := FALSE;
            tmp_CurrentStep   := ArmStep.Idle;
        END_IF;
    ELSE
        tmp_CycleDoneTimer(IN := FALSE, PT := T#0s);
    END_IF;

    IF tmp_StartTrigger THEN
        CASE TO_INT(tmp_CurrentStep) OF
            0: tmp_CurrentStep := ArmStep.Step1;
            1: MoveDown := NOT DownLimitSwitch;
               IF DownLimitSwitch THEN
                   tmp_CurrentStep := ArmStep.Step2;
               END_IF;
            2: ActivateGrip := NOT GripLimitSwitch;
               IF GripLimitSwitch THEN
                   tmp_CurrentStep := ArmStep.Step3;
               END_IF;
            3: MoveUp := NOT UpLimitSwitch;
               IF UpLimitSwitch THEN
                   tmp_CurrentStep := ArmStep.Step4;
               END_IF;
            4: MoveRight := NOT RightLimitSwitch;
               IF RightLimitSwitch THEN
                   tmp_CurrentStep := ArmStep.Step5;
               END_IF;
            5: MoveDown := NOT DownLimitSwitch;
               IF DownLimitSwitch THEN
                   tmp_CurrentStep := ArmStep.Step6;
               END_IF;
            6: ActivateRelease := NOT ReleaseLimitSwitch;
               IF ReleaseLimitSwitch THEN
                   tmp_CurrentStep := ArmStep.Step7;
               END_IF;
            7: MoveUp := NOT UpLimitSwitch;
               IF UpLimitSwitch THEN
                   tmp_CurrentStep := ArmStep.Step8;
               END_IF;
            8: MoveLeft := NOT LeftLimitSwitch;
               IF LeftLimitSwitch THEN
                   tmp_CurrentStep := ArmStep.Idle;
               END_IF;
        END_CASE;
    END_IF;

ELSIF ContinuousMode THEN
    // Same as single cycle but restarts automatically after PT delay at home
    IF Start AND NOT tmp_Gripping AND NOT tmp_Releasing THEN
        tmp_StartTrigger := TRUE;
    END_IF;

    IF tmp_CurrentStep = ArmStep.Step8 AND UpLimitSwitch AND LeftLimitSwitch THEN
        tmp_CycleDoneTimer(IN := tmp_CycleDoneTimer.Q, PT := T#1ms);
        IF tmp_CycleDoneTimer.Q THEN
            tmp_CurrentStep := ArmStep.Idle;
        END_IF;
        IF NOT tmp_CycleDoneTimer.Q AND tmp_CurrentStep = ArmStep.Idle THEN
            tmp_StartTrigger := Start;
            tmp_Gripping     := FALSE;
            tmp_Releasing    := FALSE;
        END_IF;
    ELSE
        tmp_CycleDoneTimer(IN := FALSE, PT := T#0s);
    END_IF;

    IF tmp_StartTrigger THEN
        CASE TO_INT(tmp_CurrentStep) OF
            0: tmp_CurrentStep := ArmStep.Step1;
            1: MoveDown := NOT DownLimitSwitch;
               IF DownLimitSwitch THEN
                   tmp_CurrentStep := ArmStep.Step2;
               END_IF;
            2: ActivateGrip := NOT GripLimitSwitch;
               IF GripLimitSwitch THEN
                   tmp_CurrentStep := ArmStep.Step3;
               END_IF;
            3: MoveUp := NOT UpLimitSwitch;
               IF UpLimitSwitch THEN
                   tmp_CurrentStep := ArmStep.Step4;
               END_IF;
            4: MoveRight := NOT RightLimitSwitch;
               IF RightLimitSwitch THEN
                   tmp_CurrentStep := ArmStep.Step5;
               END_IF;
            5: MoveDown := NOT DownLimitSwitch;
               IF DownLimitSwitch THEN
                   tmp_CurrentStep := ArmStep.Step6;
               END_IF;
            6: ActivateRelease := NOT ReleaseLimitSwitch;
               IF ReleaseLimitSwitch THEN
                   tmp_CurrentStep := ArmStep.Step7;
               END_IF;
            7: MoveUp := NOT UpLimitSwitch;
               IF UpLimitSwitch THEN
                   tmp_CurrentStep := ArmStep.Step8;
               END_IF;
            8: MoveLeft := NOT LeftLimitSwitch;
               IF LeftLimitSwitch THEN
                   tmp_CurrentStep := ArmStep.Idle;
               END_IF;
        END_CASE;
    END_IF;
END_IF;

END_FUNCTION_BLOCK
